# EPICS autosave request: 1.5.0/debian-12/7.0.10/modules/ADCore-ee039d2/db/NDAttribute_settings.req
file "NDTimeSeries_settings.req", P=$(P), R=$(R)TS:
file "NDPluginBase_settings.req", P=$(P), R=$(R)
